// TIA Portal project "OTOMATIK ETIKETLEME VE KUTULAMA UYGULMASI" (V18)

(* hardware
DEVICE "S7-1200 station_1"  S7-1200 Station
   slot 0: "Rack_0"  S7-1200 Rack  Rack  V1.0
   slot 1: "PLC_1"  CPU 1214C AC/DC/Rly  6ES7 214-1BG40-0XB0  V4.6
*)

// ===== PLC "PLC_1"  CPU 1214C AC/DC/Rly =====

VAR_GLOBAL   // PLC tag table "Default tag table"
   "START BUT" AT %I0.0 : Bool;
   "STOP BUT" AT %I0.1 : Bool;
   "YUKARI PISTON SEN" AT %I0.2 : Bool;
   "ASAGI PISTON SEN" AT %I0.3 : Bool;
   "ILERI PISTON SEN" AT %I0.4 : Bool;
   "GERI PISTON SEN" AT %I0.5 : Bool;
   "VALF ASAGI" AT %Q0.0 : Bool;
   "VALF YUKARI" AT %Q0.1 : Bool;
   "VALF ILERI" AT %Q0.2 : Bool;
   "START MEM" AT %M10.0 : Bool;
   "BASKI MEM" AT %M10.1 : Bool;
END_VAR

// folder: System blocks/Program resources

DATA_BLOCK "TIMER 1"   // DB1
{ S7_Optimized_Access := 'TRUE' }
AUTHOR : Simatic
FAMILY : IEC
NAME : IEC_TMR
VERSION : 1.0
// stored: InstanceOfName IEC_TIMER
"IEC_TIMER"
BEGIN
END_DATA_BLOCK

// folder: (top level)

ORGANIZATION_BLOCK "Main"   // OB1, LAD, ProgramCycle
TITLE = "Main Program Sweep (Cycle)"
{ S7_Optimized_Access := 'TRUE' }
VERSION : 0.1
   VAR_INPUT
      Initial_Call : Bool;   // Initial call of this OB
      Remanence : Bool;   // =True, if remanent data are available
   END_VAR
BEGIN

REGION Network 1: SISTEM GENEL START
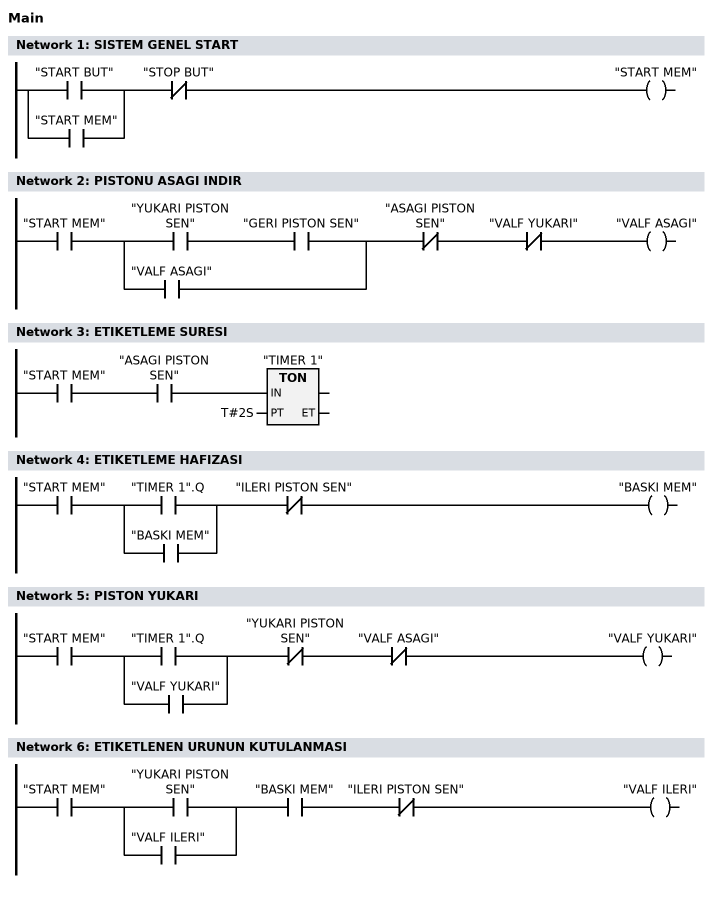
   RUNG wire#powerrail
      Contact( "START BUT" )
      wire#w1
      I_Contact( "STOP BUT" )
      Coil( "START MEM" )
   END_RUNG
   RUNG wire#powerrail
      Contact( "START MEM" )
   END_RUNG wire#w1
   // the same network as SCL:
   "START MEM" := ("START BUT" OR "START MEM") AND NOT "STOP BUT";
END_REGION

REGION Network 2: PISTONU ASAGI INDIR
   RUNG wire#powerrail
      Contact( "START MEM" )
      wire#w1
      Contact( "YUKARI PISTON SEN" )
      Contact( "GERI PISTON SEN" )
      wire#w2
      I_Contact( "ASAGI PISTON SEN" )
      I_Contact( "VALF YUKARI" )
      Coil( "VALF ASAGI" )
   END_RUNG
   RUNG wire#w1
      Contact( "VALF ASAGI" )
   END_RUNG wire#w2
   // the same network as SCL:
   "VALF ASAGI" := "START MEM" AND (("YUKARI PISTON SEN" AND "GERI PISTON SEN") OR "VALF ASAGI") AND NOT "ASAGI PISTON SEN" AND NOT "VALF YUKARI";
END_REGION

REGION Network 3: ETIKETLEME SURESI
   "TIMER 1".TON(IN := "START MEM" AND "ASAGI PISTON SEN", PT := T#2S);
END_REGION

REGION Network 4: ETIKETLEME HAFIZASI
   RUNG wire#powerrail
      Contact( "START MEM" )
      wire#w1
      Contact( "TIMER 1".Q )
      wire#w2
      I_Contact( "ILERI PISTON SEN" )
      Coil( "BASKI MEM" )
   END_RUNG
   RUNG wire#w1
      Contact( "BASKI MEM" )
   END_RUNG wire#w2
   // the same network as SCL:
   "BASKI MEM" := "START MEM" AND ("TIMER 1".Q OR "BASKI MEM") AND NOT "ILERI PISTON SEN";
END_REGION

REGION Network 5: PISTON YUKARI
   RUNG wire#powerrail
      Contact( "START MEM" )
      wire#w1
      Contact( "TIMER 1".Q )
      wire#w2
      I_Contact( "YUKARI PISTON SEN" )
      I_Contact( "VALF ASAGI" )
      Coil( "VALF YUKARI" )
   END_RUNG
   RUNG wire#w1
      Contact( "VALF YUKARI" )
   END_RUNG wire#w2
   // the same network as SCL:
   "VALF YUKARI" := "START MEM" AND ("TIMER 1".Q OR "VALF YUKARI") AND NOT "YUKARI PISTON SEN" AND NOT "VALF ASAGI";
END_REGION

REGION Network 6: ETIKETLENEN URUNUN KUTULANMASI
   RUNG wire#powerrail
      Contact( "START MEM" )
      wire#w1
      Contact( "YUKARI PISTON SEN" )
      wire#w2
      Contact( "BASKI MEM" )
      I_Contact( "ILERI PISTON SEN" )
      Coil( "VALF ILERI" )
   END_RUNG
   RUNG wire#w1
      Contact( "VALF ILERI" )
   END_RUNG wire#w2
   // the same network as SCL:
   "VALF ILERI" := "START MEM" AND ("YUKARI PISTON SEN" OR "VALF ILERI") AND "BASKI MEM" AND NOT "ILERI PISTON SEN";
END_REGION
END_ORGANIZATION_BLOCK